// TIA Portal V21 export
// export: Created 2026-11-21T13:00:31.7666517Z, ExportSetting WithDefaults, DisplayName Totally Integrated Automation Portal, DisplayVersion V21, DisplayName STEP 7 Professional, DisplayVersion V21, DisplayName STEP 7 Safety, DisplayVersion V21, DisplayName Tech WebApplication, DisplayVersion V21, DisplayName WinCC Basic/Comfort/Advanced, DisplayVersion V21, DisplayName WinCC Unified, DisplayVersion V21
VAR_GLOBAL   // PLC tag table "IO"
   Start AT %I0.0 : Bool;   // Start button
   Stop AT %I0.1 : Bool;   // Stop button, normally closed
   DoorClosed AT %I0.2 : Bool;   // Door switch
   Level AT %IW2 : Int;   // Tank level in percent
   Motor AT %Q0.0 : Bool;   // Motor contactor
   Lamp AT %Q0.1 : Bool;   // Signal lamp
   Valve AT %Q0.2 : Bool;   // Inlet valve
   Fault AT %M0.0 : Bool;   // Collected fault
   StartEdge AT %M0.1 : Bool;   // Edge memory of Start
   Setpoint AT %MW10 : Int;   // Level setpoint
   Parts AT %MW12 : Int;   // Parts counted
   Speed AT %MD20 : Real;   // Conveyor speed
   StatusWord AT %MW30 : Word;   // Status bits
   Alarm AT %M1.0 : Bool;   // Set by the sealed block
END_VAR
